Fanuc KAREL source: KB00193.KL

PROGRAM KB00193
%NOLOCKGROUP
%ENVIRONMENT MULTI
VAR
  P1: INTEGER
  P2: INTEGER
BEGIN
  P1 = 1
  P2 = 1
  UNLOCK_GROUP(P1, P2)
END KB00193
